TYPE ST_RoadParameter :
STRUCT
	nSysType: UINT;
	fRoadLenth: LREAL;
	aRoad: ARRAY[1..GVL_MC.cRoadNum] OF ST_Road;
END_STRUCT
END_TYPE

(* stored: Version 1.1.0.1, ProductVersion 3.1.4024.12
   DUT ST_RoadParameter: Id {4f1cf378-abb8-4f89-98df-74dd8db68256} *)
